(* IEC 61131-3 sources: plc-iiot-stack/src/POUs/Iiot/F_IiotIsCmdId, 2 files *)

(* ---- F_IiotIsCmdId.decl.st ---- *)
// Назначение: cmd_id по схеме: [A-Za-z0-9_-]{8,36}.
// Автор:      kr0nsch
// Версия:     0.1.0
// Документ:   docs/plc_mqtt.md, раздел «Команды»
FUNCTION F_IiotIsCmdId : BOOL
VAR_INPUT
    sText : STRING(GVL_Const.JSON_STR_LEN);
END_VAR
VAR
    iLen : INT;
    iIdx : INT;
    bCh : BYTE;
END_VAR

(* ---- F_IiotIsCmdId.impl.st ---- *)
iLen := LEN(sText);
IF iLen < UINT_TO_INT(GVL_Const.CMD_ID_MIN_LEN) OR iLen > UINT_TO_INT(GVL_Const.CMD_ID_LEN) THEN
    RETURN;
END_IF
FOR iIdx := 0 TO iLen - 1 DO
    bCh := sText[iIdx];
    IF NOT ((bCh >= GVL_Const.ASCII_UPPER_A AND bCh <= GVL_Const.ASCII_UPPER_Z)
            OR (bCh >= GVL_Const.ASCII_LOWER_A AND bCh <= GVL_Const.ASCII_LOWER_Z)
            OR (bCh >= GVL_Const.ASCII_ZERO AND bCh <= GVL_Const.ASCII_NINE)
            OR bCh = GVL_Const.ASCII_UNDERSCORE OR bCh = GVL_Const.ASCII_MINUS) THEN
        RETURN;
    END_IF
END_FOR
F_IiotIsCmdId := TRUE;
